(* IEC 61131-3 sources: plc-vscode/tests/st/all/trust-platform/crates/trust-runtime/tests/fixtures/plcopen_motion/single_axis_negative_power_enable_split/src, 2 files *)

(* ---- main.st ---- *)
PROGRAM Main
VAR
    Axis : AXIS_REF;
    Power : MC_Power;
END_VAR

Power(Axis := Axis, Enable := TRUE, EnablePositive := TRUE);
END_PROGRAM

(* ---- tests.st ---- *)
TEST_PROGRAM plcopen_motion_single_axis_negative_power_enable_split
VAR
    Axis : AXIS_REF;
    Power : MC_Power;
END_VAR

Power(Axis := Axis, Enable := TRUE, EnableNegative := TRUE);
END_TEST_PROGRAM
